TYPE ST_Channel :
STRUCT
	bActive				AT %Q*  : BOOL	 := FALSE;	
	nBrightness			AT %Q*	: UINT	 := 100; 
END_STRUCT
END_TYPE

(* stored: Version 1.1.0.1, ProductVersion 3.1.4024.12
   DUT ST_Channel: Id {ba1c87e9-366e-42cc-b50f-fb2ef855e620} *)
